// TIA Portal V21 export
// export: Created 2026-11-07T17:04:59.4445948Z, ExportSetting WithDefaults, DisplayName Totally Integrated Automation Portal, DisplayVersion V21, DisplayName STEP 7 Professional, DisplayVersion V21, DisplayName STEP 7 Safety, DisplayVersion V21, DisplayName Tech WebApplication, DisplayVersion V21, DisplayName WinCC Basic/Comfort/Advanced, DisplayVersion V21, DisplayName WinCC Unified, DisplayVersion V21
TextList "TL_Phase"  ListRange=Decimal
  TextListEntry   EntryType=SingleValue, Text="vožnja do izvora"
  TextListEntry   EntryType=SingleValue, From=1, To=1, Text="podizanje"
  TextListEntry   EntryType=SingleValue, From=2, To=2, Text="vožnja do odredišta"
  TextListEntry   EntryType=SingleValue, From=3, To=3, Text="spuštanje"
